Fanuc KAREL source: kb00078.KL

-- PROVISIONAL review KL for V1013-1; original PC SHA256 3213fe41140515e2b307039ec37992d28630b9b22ffcd534fd4fc6c1cc2f78b3
-- Incomplete behavior may be omitted. Consult companion uncertainty JSON. Do not deploy.
PROGRAM KB00078
%NOLOCKGROUP
BEGIN
  -- UNRESOLVED_PC offsets 5-21; opcodes 27,22,31,23
  -- UNRESOLVED_PC offsets 26-30; opcodes 7F
END KB00078
